// TIA Portal V19 export
DATA_BLOCK "iFB_Conveyor_Test"   // DB4
// stored: InstanceOfName FB_Conveyor_Test, InstanceOfType FB
"FB_Conveyor_Test"
BEGIN
END_DATA_BLOCK
